// Generated by voz_llm_plc_agent
// Target: Siemens TIA Portal V18 - SCL external source
// Review and compile before any download to physical hardware.

FUNCTION_BLOCK "PLC_PRG"
{ S7_Optimized_Access := 'TRUE' }
VERSION : 0.1
VAR_INPUT
   I_Start : Bool := FALSE;
   I_Emergency : Bool := FALSE;
   I_Alarm_Active : Bool := FALSE;
END_VAR
VAR_OUTPUT
   Q_VFD_Enable : Bool := FALSE;
END_VAR
BEGIN
(* Habilitacion solo mientras no exista una alarma activa (condicion de entrada) *)
#Q_VFD_Enable := #I_Start AND NOT #I_Alarm_Active AND NOT #I_Emergency;
END_FUNCTION_BLOCK

DATA_BLOCK "DB_PLC_PRG"
{ S7_Optimized_Access := 'TRUE' }
VERSION : 0.1
NON_RETAIN
"PLC_PRG"
BEGIN
END_DATA_BLOCK

ORGANIZATION_BLOCK "Main"
{ S7_Optimized_Access := 'TRUE' }
VERSION : 0.1
BEGIN
   "DB_PLC_PRG"(
      I_Start := "I_Start",
      I_Emergency := "I_Emergency",
      I_Alarm_Active := "I_Alarm_Active",
      Q_VFD_Enable => "Q_VFD_Enable"
   );
END_ORGANIZATION_BLOCK
